TYPE ST_Cia402Config :
STRUCT
    tStateTimeout     : TIME := T#2S;     // each transition, the mode switch
    tStopTimeout      : TIME := T#10S;    // a step down, a fault reaction
    tHomingTimeout    : TIME := T#60S;    // one whole homing run
    nResetAttempts    : UINT := 3;        // fault resets; 0 counts as 1
    tResetPause       : TIME := T#1S;     // between two reset attempts
    bQuickStopStays   : BOOL := FALSE;    // 0x605A is 5-8 on this drive
    nStandstillWindow : DINT := 0;        // position band, 0x6064 units
    tStandstill       : TIME := T#100MS;  // in the band this long: stopped
    tInputsInvalid    : TIME := T#100MS;  // bInputsValid FALSE this long: error
    bEnableAfterReset : BOOL := FALSE;    // TRUE: re-enable after bReset, as MC_Power
END_STRUCT
END_TYPE

(* stored: Version 1.1.0.1, ProductVersion 3.1.4024.0
   DUT ST_Cia402Config: Id {70c0f2f9-addd-4b57-bccd-dc623a854d93} *)
